(* PLC project g_building_lighting_clean, Anonymous Benchmark Suite 1.0 *)
(* stored: creationDateTime 2026-07-09T00:00:00 *)

PROGRAM g_building_lighting_clean
  VAR_INPUT
    demand : BOOL;
    master_off : BOOL;
    maint : BOOL;
  END_VAR
  VAR_OUTPUT
    lights : BOOL;
    setback : BOOL;
  END_VAR

(* LD diagram, written out as Structured Text *)
lights := NOT master_off AND demand;
setback := master_off;
END_PROGRAM

CONFIGURATION Config0
  RESOURCE Res0 ON PLC
    TASK tcyclic(INTERVAL := T#10ms, PRIORITY := 0);
    PROGRAM inst0 WITH tcyclic : g_building_lighting_clean;
  END_RESOURCE
END_CONFIGURATION
